Fanuc KAREL source: KX00030.KL

PROGRAM KX00030
%NOLOCKGROUP
%NOPAUSE = ERROR + COMMAND
VAR
  I: INTEGER
  J: INTEGER
  B: BOOLEAN
  F: FILE
  S: STRING[80]
  P: XYZWPR
BEGIN
  I = 1
END KX00030
